(* IEC 61131-3 sources: tsplc/examples/bottling-line/raw-st/src/capping/FB_Capper, 2 files *)

(* ---- declaration.st ---- *)
FUNCTION_BLOCK FB_Capper
VAR_INPUT
	BottlePresent : BOOL;
END_VAR
VAR_OUTPUT
	Running : BOOL;
END_VAR
VAR
	State : E_CapperState := E_CapperState.Idle;
	Capped : UDINT;
END_VAR

(* ---- FB_Capper.implementation.st ---- *)
CASE State OF
	E_CapperState.Idle:
		IF BottlePresent THEN
			State := E_CapperState.Capping;
		END_IF
	E_CapperState.Capping:
		Capped := Capped + 1;
		State := E_CapperState.Idle;
END_CASE
Running := State = E_CapperState.Capping;
